TYPE HmiStatus :
STRUCT
	acknowledgedSequence : UDINT;
	missionState : MissionState;
	lastRejection : STRING(80);
	estimatedPose : Pose2D;
	isSimulatorConnected : BOOL;
	isLidarOk : BOOL;
	hasMap : BOOL;
END_STRUCT
END_TYPE

(* stored: Version 1.1.0.1, ProductVersion 3.1.4026.12
   DUT HmiStatus: Id {6dc03ffe-a80b-54c4-a7a6-fbb20cd05687} *)
